(* PLC project probe.project, CODESYS CODESYS V3.5 SP17 Patch 3 *)
(* stored: creationDateTime 2026-10-20T03:54:26.7214605, modificationDateTime 1601-01-01T03:00:00 *)

TYPE E_ProbeMode : (Off := 0, Manual := 1, Auto := 2);
END_TYPE
